(* IEC 61131-3 sources: ConveyorControl-with-PLC/4E_Gruppe1_Graf_Projekt1_HMI/Network/LseRtkMain, 1 file *)

(* ---- ONE_LseRtkMain_Table.st ---- *)
#define OBJECTS_CONFIG

//Define part of class KeyPadNum
#define NUMBUT_WIDTH   60
#define NUMBUT_HEIGHT  50
#define NUMBUT_XOFF     6
#define NUMBUT_YOFF   100
#define NUMPAD_WIDTH  251
#define NUMPAD_HEIGHT 305

FUNCTION GLOBAL TAB ONE_LseRtkMain
-1$UINT, 0$UINT,
0$UINT, 0$UINT,

9$UDINT,
TO_UDINT(3788417926), "_Global", 0$UINT, 12$UINT, 0$UINT,
TO_UDINT(1552551876), "_Lse", 0$UINT, 101$UINT, 1$UINT,
TO_UDINT(3599188277), "_Screen", 0$UINT, 2$UINT, 0$UINT,
TO_UDINT(3931827689), "_SysDateTime", 0$UINT, 5$UINT, 1$UINT,
TO_UDINT(3192771746), "_XAccess", 0$UINT, 1$UINT, 1$UINT,
TO_UDINT(2266234845), "KeyPadAnum", 0$UINT, 6$UINT, 1$UINT,
TO_UDINT(1581172638), "KeyPadImages", 0$UINT, 1$UINT, 2$UINT,
TO_UDINT(2771413771), "KeyPadNum", 0$UINT, 3$UINT, 1$UINT,
TO_UDINT(1903583397), "Ram", 1$UINT, 3$UINT, 5$UINT,

_NO_ATTR, TO_UDINT(299963966), "LSE",

_NO_ATTR, TO_UDINT(3035062039), "SYSDATETIME",

_NO_ATTR, TO_UDINT(3799848273), "XACCESS0",

_NO_ATTR, TO_UDINT(2266234845), "KEYPADANUM",

1$UINT, TO_UDINT(943717585), "KEYPADANUM\KEYPADIMG",
1$UINT, TO_UDINT(3532807661), "KEYPADNUM\KEYPADIMG",

_NO_ATTR, TO_UDINT(2771413771), "KEYPADNUM",

1$UINT, TO_UDINT(1119588755), "SYSDATETIME\SUMMERTIME",
1$UINT, TO_UDINT(440852310), "XACCESS0\RAM0",
1$UINT, TO_UDINT(1833037760), "XACCESS0\RAM1",
1$UINT, TO_UDINT(4098408058), "XACCESS0\RAM2",
1$UINT, TO_UDINT(2203029228), "XACCESS0\RAM3",

//Internal connections
0$UDINT,
7$UDINT,
TO_UDINT(1), "SummerTime", TO_UDINT(7),
TO_UDINT(2), "Ram0", TO_UDINT(8),
TO_UDINT(2), "Ram1", TO_UDINT(9),
TO_UDINT(2), "Ram2", TO_UDINT(10),
TO_UDINT(2), "Ram3", TO_UDINT(11),
TO_UDINT(3), "KeyPadImg", TO_UDINT(4),
TO_UDINT(6), "KeyPadImg", TO_UDINT(5),
0$UDINT,
3$UDINT,
TO_UDINT(2), "Lse", TO_UDINT(0), "Lse",
TO_UDINT(3), "Lse", TO_UDINT(0), "Lse",
TO_UDINT(6), "Lse", TO_UDINT(0), "Lse",

//Initialization values
0$UDINT,
9$UDINT,
TO_UDINT(0), "AmericanDateFormat", TO_UDINT(0),//|LseRtkMain.Lse.AmericanDateFormat;
TO_UDINT(0), "SeekAlgorithm", TO_UDINT(1),//|LseRtkMain.Lse.SeekAlgorithm;
TO_UDINT(1), "DoSummerTime", TO_UDINT(0),//|LseRtkMain.SysDateTime.DoSummerTime;
TO_UDINT(3), "No", TO_UDINT(_WIN_EDITOR_ANUMERIC),//|LseRtkMain.KeyPadAnum.No;
TO_UDINT(3), "ImA", TO_UDINT(IMA_WINDOW),//|LseRtkMain.KeyPadAnum.ImA;
TO_UDINT(3), "AltGr", TO_UDINT(1),//|LseRtkMain.KeyPadAnum.AltGr;
TO_UDINT(3), "CapitalLetter", TO_UDINT(0),//|LseRtkMain.KeyPadAnum.CapitalLetter;
TO_UDINT(6), "No", TO_UDINT(_WIN_EDITOR_NUMERIC),//|LseRtkMain.KeyPadNum.No;
TO_UDINT(6), "ImA", TO_UDINT(IMA_WINDOW),//|LseRtkMain.KeyPadNum.ImA;

//Symbolic initialization values
0$UDINT,
0$UDINT,

//Initialization of string values
0$UDINT,
0$UDINT,

//Configuration of tasks (RealTime, Cyclic, Background)
0$UDINT,
0$UDINT,

0$UDINT,
0$UDINT,

0$UDINT,
2$UDINT,
TO_UDINT(0), (-1)$UDINT, 4194303$DINT, 	//LSE
TO_UDINT(1), (100)$UDINT, 4194303$DINT, 	//SYSDATETIME

//External connections
0$UDINT,
0$UDINT,

//Magic internal connections
0$UDINT,
0$UDINT,

//Configuration of timeslots of tasks (RealTime, Cyclic)
#ifdef __LSLLDR_TIMESLOTS__
0$UDINT,
0$UDINT,

0$UDINT,
0$UDINT,

#endif //__LSLLDR_TIMESLOTS__

//MultiMaster connections
#ifdef __LSLLDR_MULTIMASTER__
0$UDINT,
0$UDINT,
#endif //__LSLLDR_MULTIMASTER__

END_FUNCTION
